(* IEC 61131-3 sources: model-first-plc-agent-ai/results/T2-W-06, 2 files *)

(* ---- a1_code.st ---- *)
FUNCTION_BLOCK FillingRuntime
VAR_INPUT
    start : BOOL;
    stop : BOOL;
    LSH : BOOL;
    LSHH : BOOL;
    TimerDuration : TIME;
END_VAR
VAR_OUTPUT
    fill_valve : BOOL;
    discharge_valve : BOOL;
END_VAR
VAR
    x0 : BOOL := TRUE;
    x1 : BOOL := FALSE;
    previous_x1 : BOOL;
    timer_done : BOOL := FALSE;
    filling_timer : TON;
END_VAR

(* Evaluate elapsed time for the currently active step. *)
filling_timer(IN := x1, PT := TimerDuration);
timer_done := filling_timer.Q;
previous_x1 := x1;

(* Evaluate transitions from the current situation. *)
IF x0 THEN
    IF start AND NOT stop AND NOT LSHH THEN
        x0 := FALSE;
        x1 := TRUE;
    END_IF;
ELSIF x1 THEN
    IF stop OR LSHH OR timer_done THEN
        x1 := FALSE;
        x0 := TRUE;
    END_IF;
END_IF;

(* Start timing on entry and reset timing on exit. *)
IF x1 <> previous_x1 THEN
    filling_timer(IN := x1, PT := TimerDuration);
    timer_done := FALSE;
END_IF;

fill_valve := x1;
discharge_valve := FALSE;

END_FUNCTION_BLOCK

PROGRAM Main
VAR
    StartCommand AT %IX100.0 : BOOL;
    StopCommand AT %IX100.1 : BOOL;
    LSH AT %IX100.2 : BOOL;
    LSHH AT %IX100.3 : BOOL;
    FillValve AT %QX100.0 : BOOL;
    DischargeValve AT %QX100.1 : BOOL;
END_VAR
VAR
    TimerDuration : TIME := T#0s;
    start_edge : R_TRIG;
    filling_control : FillingRuntime;
END_VAR

(* Initialization is provided by the declared initial values. *)
start_edge(CLK := StartCommand);

filling_control(
    start := start_edge.Q,
    stop := StopCommand,
    LSH := LSH,
    LSHH := LSHH,
    TimerDuration := TimerDuration
);

FillValve := filling_control.fill_valve;
DischargeValve := filling_control.discharge_valve;

END_PROGRAM

(* ---- a2_code.st ---- *)
FUNCTION_BLOCK FB_TimedTankFilling
VAR_INPUT
    StartCommand : BOOL;
    StopCommand : BOOL;
    LSH : BOOL;
    LSHH : BOOL;
    TimerDuration : TIME;
END_VAR
VAR_OUTPUT
    FillValve : BOOL;
    DischargeValve : BOOL;
END_VAR
VAR
    StartEdge : R_TRIG;
    FillingTimer : TON;
    ActiveState : INT := 0;
    start : BOOL;
    stop : BOOL;
    timer_done : BOOL;
    fill_valve : BOOL;
    discharge_valve : BOOL;
END_VAR

StartEdge(CLK := StartCommand);
start := StartEdge.Q;
stop := StopCommand;

IF stop THEN
    ActiveState := 0;
ELSE
    CASE ActiveState OF
        0:
            IF start THEN
                ActiveState := 1;
            END_IF;
        1:
            ActiveState := 1;
    ELSE
        ActiveState := 0;
    END_CASE;
END_IF;

FillingTimer(
    IN := (ActiveState = 1),
    PT := TimerDuration
);
timer_done := FillingTimer.Q;

IF ActiveState = 1 THEN
    IF stop OR timer_done OR LSHH THEN
        ActiveState := 0;
    END_IF;
END_IF;

IF ActiveState = 0 THEN
    FillingTimer(IN := FALSE, PT := TimerDuration);
    timer_done := FALSE;
END_IF;

fill_valve := (ActiveState = 1);
discharge_valve := FALSE;

FillValve := fill_valve;
DischargeValve := discharge_valve;

END_FUNCTION_BLOCK

PROGRAM Main
VAR
    StartCommand AT %IX100.0 : BOOL;
    StopCommand AT %IX100.1 : BOOL;
    LSH AT %IX100.2 : BOOL;
    LSHH AT %IX100.3 : BOOL;
    FillValve AT %QX100.0 : BOOL;
    DischargeValve AT %QX100.1 : BOOL;
END_VAR
VAR
    TimerDuration : TIME;
    TankController : FB_TimedTankFilling;
END_VAR

TankController(
    StartCommand := StartCommand,
    StopCommand := StopCommand,
    LSH := LSH,
    LSHH := LSHH,
    TimerDuration := TimerDuration
);

FillValve := TankController.FillValve;
DischargeValve := TankController.DischargeValve;

END_PROGRAM
